TYPE ST_DosingStationConfiguration :
STRUCT
	ratio				: LREAL := 0.2; //dosing flow / main flow while running
END_STRUCT
END_TYPE

(* stored: Version 1.1.0.1, ProductVersion 3.1.4024.12
   DUT ST_DosingStationConfiguration: Id {4c75bb2e-06d8-441d-8788-4fd2b9203f7f} *)
